// TIA Portal V20 export
TYPE "WT2_Vr_Status_UDT"
   STRUCT
      iHandshake : Int;
      Fehler : Struct
         bE0000_KonfigFehler : Bool;
         bE0001_Reserviert : Bool;
         bE0002_InvUngueltig : Bool;
         bE0003_Reserviert : Bool;
         bE0004_FrostschutzFehler : Bool;
         bE0005_VrPumpeFehlerBetr : Bool;
         bE0006_VrPumpeFehlerStillstand : Bool;
         bE0007_VrEintrittWarm : Bool;
         bE0008_NivAbschHochFehler : Bool;
         bE0009_KonfigFehlerUmstDIPol : Bool;
         bE0010_Reserviert : Bool;
         bE0011_Reserviert : Bool;
         bE0012_NivAbsch2HochFehler : Bool;
         bE0013_KonfigFehlerOelrekt : Bool;
         bE0014_Resreviert : Bool;
         bE0015_Reserviert : Bool;
         bE0016_MedUeberdruckZuTief : Bool;
         b041_Reserve : Bool;
         b042_Reserve : Bool;
         b043_Reserve : Bool;
         b044_Reserve : Bool;
         b045_Reserve : Bool;
         b046_Reserve : Bool;
         b047_Reserve : Bool;
         by05_Reserve : Byte;
      END_STRUCT;
      Alarm : Struct
         bA1000_Reserviert : Bool;
         bA1001_SlaveAusgef : Bool;
         bA1002_Reserviert : Bool;
         bA1003_HauptMasterAusgef : Bool;
         bA1004_Reserviert : Bool;
         bA1005_Reserviert : Bool;
         bA1006_Reserviert : Bool;
         bA1007_Reserviert : Bool;
         bA1008_Reserviert : Bool;
         bA1009_Reserviert : Bool;
         bA1010_MVrMasterAktiv : Bool;
         bA1011_ObjektIDMehrfVorhanden : Bool;
         bA1012_Reserviert : Bool;
         bA1013_Reserviert : Bool;
         bA1014_AlarmNivAbschEndsch : Bool;
         bA1015_AlarmNivAbsch2Endsch : Bool;
         bA1016_Reserviert : Bool;
         b081_Reserve : Bool;
         b082_Reserve : Bool;
         b083_Reserve : Bool;
         b084_Reserve : Bool;
         b085_Reserve : Bool;
         b086_Reserve : Bool;
         b087_Reserve : Bool;
         by09_Reserve : Byte;
      END_STRUCT;
      Zustand : Struct
         bFehlerzustandAktiv : Bool;
         bAlarmzustandAktiv : Bool;
         bSystemMeldungAktiv : Bool;
         bSeviceMeldungAktiv : Bool;
         bStopManuell : Bool;
         bStopAuto : Bool;
         bStopExtern : Bool;
         bBetriebAuto : Bool;
         bBetriebManuell : Bool;
         bAnlaufAuto : Bool;
         bAnlaufManuell : Bool;
         bManuellStoppen : Bool;
         b114_Reserve : Bool;
         b115_Reserve : Bool;
         b116_Reserve : Bool;
         b117_Reserve : Bool;
         by12_Reserve : Byte;
         bInventarAufnahme : Bool;
         b131_Reserve : Bool;
         bStandbyMasterInit : Bool;
         bStandbyMasterPassiv : Bool;
         bStandbyMasterAktiv : Bool;
         bMasterGesperrt : Bool;
         bSollwertAbsenkung : Bool;
         b137_Reserve : Bool;
         by14_Reserve : Byte;
         by15_Reserve : Byte;
         by16_Reserve : Byte;
         by17_Reserve : Byte;
      END_STRUCT;
      DigIn : Struct
         bSollwertB : Bool;
         bRMVrPumpe : Bool;
         bTKSDigital : Bool;
         bStartbefehlKS : Bool;
         bAbschNivHoch : Bool;
         bAbschNiveauregFreigabe : Bool;
         bAbsch2NivHoch : Bool;
         bAbsch2NiveauregFreigabe : Bool;
         bAbschBetriebsart : Bool;
         bAbsch2Betriebsart : Bool;
         bAbschNivEndschOffen : Bool;
         bAbschNivEndschGeschl : Bool;
         bAbsch2NivEndschOffen : Bool;
         bAbsch2NivEndschGeschl : Bool;
         bFrostschutzDigital : Bool;
         bMediumKreislUeberdruck : Bool;
         by20_Reserve : Byte;
         by21_Reserve : Byte;
      END_STRUCT;
      DigOut : Struct
         bStartbefehlVrPumpe : Bool;
         bMVKS : Bool;
         bAbschNiveaureg : Bool;
         bAbsch2Niveaureg : Bool;
         bMVAbschNachspeisung : Bool;
         bMVAbsch2Nachspeisung : Bool;
         bOelrektifizierung : Bool;
         b227_Reserve : Bool;
         by23_Reserve : Byte;
         by24_Reserve : Byte;
         by25_Reserve : Byte;
      END_STRUCT;
      chReserve1 : Char;
      chVrReglerEinheit : Char;
      rVrRegIst : Real;
      rVrRegSoll : Real;
      rVrRegOut : Real;
      rVrTempEintritt : Real;
      rVrTempAustritt : Real;
      rReserveReal : Array[0..3] of Real;
   END_STRUCT;
END_TYPE
